(* IEC 61131-3 sources: volt/packages/volt-lsp-iec/test-corpus/lenze-mid/Device/Plc Logic/Application/Library Manager/L_IMHP_ModuleHandler, 81 files *)

(* ---- L_IMHP_COMPONENTTYPE.dut ---- *)
TYPE L_IMHP_COMPONENTTYPE :
(
	DEVICE := 101,
	IEC_RUNTIME := 102,
	LINUX_RUNTIME := 103,
	FAST_UI_RUNTIME := 104,
	FRAMEWORKSERVICE := 105,
	DEVICEFEATURES := 106,
	ETHERCATSLAVE := 201,
	ETHERCATMASTER := 202,
	FIELDBUSSLAVE := 203,
	FIELDBUSMASTER := 204,
	ETHERNET := 205,
	OPC_UA_CLIENT := 206,
	OPC_UA_SERVER := 207,
	UI_CLIENT := 208,
	UI_SERVER := 209,
	SINGLEAXISKINEMATICS := 301,
	SINGLEAXISKINEMATIK := 301,
	ROBOTKINEMATICS := 302,
	ROBOTKINEMATIC := 302,
	LOGICAXIS := 401,
	MOTIONAXIS := 402,
	VIRTUALAXIS := 403,
	ENCODERAXIS := 404,
	VIRTUALENCODERAXIS := 405,
	TECHNOLOGYFUNCTIONS := 500,
	TECHNOLOGYMODULE := 501,
	TECHNOLOGYAPPLICATION := 503,
	MACHINEMODULE := 504,
	MOTIONBASE := 505,
	COORDINATEDMOTION := 506,
	GENERALMACHINEMODULE := 551,
	GENERALAPPLICATIONMODULE := 552,
	DATAMANAGEMENT := 601,
	CLOUDCONNECTIVITY := 602,
	DATAANALYTICS := 603
);
END_TYPE

(* ---- L_IMHP_EM_CLEARERRORDATA.dut ---- *)
TYPE L_IMHP_EM_CLEARERRORDATA :
STRUCT
	VERSION : UDINT := 1;
	WERRORID : WORD;
	WTEXTREFID : WORD;
END_STRUCT
END_TYPE

(* ---- L_IMHP_EM_COMMAND.dut ---- *)
TYPE L_IMHP_EM_COMMAND :
(
	NOCOMMAND := 0,
	NOTIFYERROR := 1,
	NOTIFYERRORSHORT := 2,
	CLEARERROR := 3,
	RESETERROR := 4
);
END_TYPE

(* ---- L_IMHP_EM_EVENTPARAMETERS.dut ---- *)
TYPE L_IMHP_EM_EVENTPARAMETERS :
STRUCT
	EVENTPARAMETERS : ARRAY [1..10] OF L_IMHP_EM_ParameterItem;
END_STRUCT
END_TYPE

(* ---- L_IMHP_EM_EVENTPARAMETERSSHORT.dut ---- *)
TYPE L_IMHP_EM_EVENTPARAMETERSSHORT :
STRUCT
	EVENTPARAMETERS : ARRAY [1..10] OF L_IMHP_EM_ParameterItemShort;
END_STRUCT
END_TYPE

(* ---- L_IMHP_EM_NOTIFYERRORDATA.dut ---- *)
TYPE L_IMHP_EM_NOTIFYERRORDATA :
STRUCT
	VERSION : UDINT := 1;
	WERRORID : WORD;
	WTEXTREFID : WORD;
	SEVERITY : USINT;
	PRIORITY : USINT;
	GROUP : USINT;
END_STRUCT
END_TYPE

(* ---- L_IMHP_EM_PARAMETERITEM.dut ---- *)
TYPE L_IMHP_EM_PARAMETERITEM :
STRUCT
	SIZE : BYTE;
	ETYPE : INT;
	VALUE : L_IMHP_EM_ParaValue;
END_STRUCT
END_TYPE

(* ---- L_IMHP_EM_PARAMETERITEMSHORT.dut ---- *)
TYPE L_IMHP_EM_PARAMETERITEMSHORT :
STRUCT
	SIZE : BYTE;
	ETYPE : INT;
	VALUE : L_IMHP_EM_ParaValueShort;
END_STRUCT
END_TYPE

(* ---- L_IMHP_EM_PARAVALUE.dut ---- *)
TYPE L_IMHP_EM_PARAVALUE :
UNION
	DWVALUE : DWORD;
	DNVALUE : DINT;
	FVALUE : REAL;
	STVALUE : STRING;
	DWTEXTLISTID : DWORD;
END_UNION
END_TYPE

(* ---- L_IMHP_EM_PARAVALUESHORT.dut ---- *)
TYPE L_IMHP_EM_PARAVALUESHORT :
UNION
	DWVALUE : DWORD;
	DNVALUE : DINT;
	RVALUE : REAL;
	LRVALUE : LREAL;
	DWTEXTLISTID : DWORD;
END_UNION
END_TYPE

(* ---- L_IMHP_EM_REGISTERDATA.dut ---- *)
TYPE L_IMHP_EM_REGISTERDATA :
STRUCT
	VERSION : UDINT := 1;
	CMPNAME : POINTER TO STRING;
	LAYER : BYTE;
	TEXTREFID : WORD;
	ADDITIONALCMPINFOS : DWORD;
END_STRUCT
END_TYPE

(* ---- L_IMHP_EM_SERVERITYLEVEL.dut ---- *)
TYPE L_IMHP_EM_SERVERITYLEVEL :
(
	NO_RESPONSE := 0,
	FAULT_CIA402 := 1,
	WARNING := 2,
	INFORMATION := 11,
	WARNING_LOCK := 13,
	TROUBLE_LOG := 15,
	TROUBLE := 16,
	FAULT_LOG := 18,
	FAULT_FAST_STOP := 19,
	FAULT_QSP := 20,
	FAULT_QSP_CINH := 21,
	FAULT := 23
);
END_TYPE

(* ---- L_IMHP_LAYER.dut ---- *)
TYPE L_IMHP_LAYER :
(
	BASE_SETTINGS := 4,
	COMMUNICATION := 5,
	KINEMATICS := 6,
	MOTION := 7,
	TECH_APPLICATION := 8,
	PROCESS_CONTROL := 9
);
END_TYPE

(* ---- L_IMHP_LM_APPLICATIONCREDITCONFIGURATION.dut ---- *)
TYPE L_IMHP_LM_APPLICATIONCREDITCONFIGURATION :
STRUCT
	VERSION : DWORD := 1;
	SIZE : DWORD := SIZEOF(L_IMHP_LM_ApplicationCreditConfiguration);
	FAST_TOOLBOX : DWORD := 0;
	FAST_SERVICES : DWORD := 0;
	FAST_UI : DWORD := 0;
	OPC_UA : DWORD := 0;
	DEVICE_FEATURES : DWORD := 0;
	ADDITIONAL_BUDGETS : ARRAY [0..14] OF DWORD := [0, 0, 0, 0, 0, 0, 0, 0, 0, 0, 0, 0, 0, 0, 0];
END_STRUCT
END_TYPE

(* ---- L_IMHP_LM_APPLICATIONCREDITINFO.dut ---- *)
TYPE L_IMHP_LM_APPLICATIONCREDITINFO :
STRUCT
	VERSION : DWORD := 1;
	SIZE : DWORD := SIZEOF(L_IMHP_LM_ApplicationCreditInfo);
	AVAILABLEAPPLICATIONCREDIT : DWORD := 0;
	MAXAPPLICATIONCREDIT : DWORD := 0;
	USEDAPPLICATIONCREDIT : DWORD := 0;
END_STRUCT
END_TYPE

(* ---- L_IMHP_LM_BLISTDATA.dut ---- *)
TYPE L_IMHP_LM_BLISTDATA :
STRUCT
	VERSION : DWORD := 1;
	SIZE : DWORD := SIZEOF(L_IMHP_LM_BListData);
	COMPONENTNAME : POINTER TO STRING := 0;
	INSTANCEPATH : POINTER TO STRING := 0;
END_STRUCT
END_TYPE

(* ---- L_IMHP_LM_COMMAND.dut ---- *)
TYPE L_IMHP_LM_COMMAND :
(
	NOCOMMAND := 0,
	WRITECOMPONENTLIST := 1,
	GETAPPCREDITOFCOMPONENT := 2,
	GETAPPCREDITINFO := 3,
	ACTIVATEAPPCREDIT := 4,
	GETMODIFICATIONTIME := 5
);
END_TYPE

(* ---- L_IMHP_LM_CONFIGMODEDATA.dut ---- *)
TYPE L_IMHP_LM_CONFIGMODEDATA :
STRUCT
	VERSION : DWORD := 1;
	SIZE : DWORD := SIZEOF(L_IMHP_LM_ConfigModeData);
	UDICONFIGMODE : UDINT := 0;
END_STRUCT
END_TYPE

(* ---- L_IMHP_LM_CONFIGURECOMMAND.dut ---- *)
TYPE L_IMHP_LM_CONFIGURECOMMAND :
(
	NOCOMMAND := 0,
	APPCREDITCONFIGURATION := 1,
	SETCONFIGMODE := 2,
	STARTONLINECHANGEHANDLING := 3,
	FINISHONLINECHANGEHANDLING := 4
);
END_TYPE

(* ---- L_IMHP_LM_LICENSCLASS.dut ---- *)
TYPE L_IMHP_LM_LICENSCLASS :
(
	T := 1,
	F := 2,
	I := 3
);
END_TYPE

(* ---- L_IMHP_LM_REGISTERDATA.dut ---- *)
TYPE L_IMHP_LM_REGISTERDATA :
STRUCT
	VERSION : DWORD := 1;
	SIZE : DWORD := SIZEOF(L_IMHP_LM_RegisterData);
	APPLICATIONCREDIT : DWORD := 0;
	LICENSECLASS : DWORD := 0;
	LICENSECLASSNUMBER : DWORD := 0;
END_STRUCT
END_TYPE

(* ---- L_IMHP_MH_COMMAND.dut ---- *)
TYPE L_IMHP_MH_COMMAND :
(
	UPDATEACTIVESTATUS := 0,
	UPDATECOMMUNICATIONADRESS := 1,
	UPDATEPARENTCHILDRELATION := 2,
	UPDATECOMPONENTTYPE := 3,
	UPDATECOMPONENTNAME := 4
);
END_TYPE

(* ---- L_IMHP_MODULEINFO.dut ---- *)
TYPE L_IMHP_MODULEINFO :
STRUCT
	DWID : DWORD;
	SNAME : STRING;
	SPATH : STRING(255);
	SCOMMPATH : STRING(199);
	ELAYER : L_IMHP_Layer := L_IMHP_Layer.Tech_Application;
	ECOMPTYPE : L_IMHP_ComponentType := L_IMHP_ComponentType.GeneralApplicationModule;
	ESUBCOMPTYPE : DWORD;
	XCOMPACTIVE : BOOL;
	WCHILDCOUNT : WORD;
	WTEXTREFID : WORD;
	XUSELEM : BOOL;
	XUSELLM : BOOL;
	RELATIONSHIPID : L_IMHP_RelationshipID := L_IMHP_RelationshipID.ApplicationView;
	PARENTMODULE : L_IMHP_IModuleHandler;
END_STRUCT
END_TYPE

(* ---- L_IMHP_RELATIONSHIPDATA.dut ---- *)
TYPE L_IMHP_RELATIONSHIPDATA :
STRUCT
	VERSION : UDINT := 1;
	SIZE : UDINT := SIZEOF(L_IMHP_RelationshipData);
	RELATIONSHIPID : L_IMHP_RelationshipID;
	PARENTHANDLE : RTS_IEC_HANDLE;
END_STRUCT
END_TYPE

(* ---- L_IMHP_RELATIONSHIPID.dut ---- *)
TYPE L_IMHP_RELATIONSHIPID :
(
	NORELATIONSHIP := 0,
	APPLICATIONVIEW := 1,
	COMMUNICATIONVIEW := 2,
	ASSETVIEW := 3
);
END_TYPE

(* ---- L_IMHP_REQUESTEDSERVICE.dut ---- *)
TYPE L_IMHP_REQUESTEDSERVICE :
STRUCT
	VERSION : UDINT := 1;
	SIZE : UDINT := SIZEOF(L_IMHP_RequestedService);
	SERVICEID : L_IMHP_ServiceID;
	SIZEOFREGISTRATIONDATA : UDINT;
	PREGISTRATIONDATA : POINTER TO BYTE;
	SERVICEAVAILABLE : UDINT;
	SERVICEVERSION : UDINT;
	REGISTRATIONSTATUS : UDINT;
	SIZEOFRESULTDATA : UDINT;
	PRESULTDATA : POINTER TO BYTE;
END_STRUCT
END_TYPE

(* ---- L_IMHP_SERVICEAVAILABLEDATA.dut ---- *)
TYPE L_IMHP_SERVICEAVAILABLEDATA :
STRUCT
	VERSION : UDINT := 1;
	SIZE : UDINT := SIZEOF(L_IMHP_ServiceAvailableData);
	SERVICEID : L_IMHP_ServiceID;
	SERVICEAVAILABLE : UDINT;
	SERVICEVERSION : UDINT;
END_STRUCT
END_TYPE

(* ---- L_IMHP_SERVICEID.dut ---- *)
TYPE L_IMHP_SERVICEID :
(
	NOSERVICE := 0,
	LENZEMODULEHANDLER := 1,
	LENZEERRORMANAGEMENT := 2,
	LENZESTATEHANDLER := 3,
	LENZELICENSEMANAGER := 4,
	LENZEASSETMANAGER := 5
);
END_TYPE

(* ---- L_IMHP_CONSTANTS.gvl ---- *)
VAR_GLOBAL
	GC_MAXCOMPIDX : WORD := 100;
END_VAR

(* ---- L_IMHP_INTERN.gvl ---- *)
VAR_GLOBAL
	XERRORHANDLINGFORI950 : BOOL;
	DEVICEMODULEHANDLER : L_IMHP_DeviceModule;
	COMPONENTREGISTRATION : L_IMHP_HandleComponentRegistration;
END_VAR

(* ---- L_IMHP_IFASTFRAMECONFIG.itf ---- *)
INTERFACE L_IMHP_IFASTFRAMECONFIG
END_INTERFACE

METHOD ADDPARAMETERINTERFACE
VAR_INPUT
	IIODRVPARAMETER : ICmpIoDrvParameter;
END_VAR
END_METHOD

(* ---- L_IMHP_IMODULEHANDLER.itf ---- *)
INTERFACE L_IMHP_IMODULEHANDLER
END_INTERFACE

METHOD ACTIVATEAPPCREDITS : BOOL
VAR_INPUT
	XACTIVATE : BOOL;
END_VAR
END_METHOD

METHOD ADDAPPCREDIT
VAR_INPUT
	CREDIT : UDINT;
END_VAR
END_METHOD

METHOD CHECKERRORRESETOCCURED : BOOL
VAR_IN_OUT
	RESETTIME : SYSTIME;
END_VAR
END_METHOD

METHOD CHECKERRORRESETTRIGGER : BOOL
VAR_IN_OUT
	LASTTRIGGERTIME : TIME;
END_VAR
END_METHOD

METHOD CLEARSEVERITYANDREACTION
VAR_INPUT
	ESEVERITY : USINT;
	DISEVERITYCOUNT : DINT;
	EREACTION : WORD;
	DIREACTIONCOUNT : DINT;
	XHANDLEASFORWARDEDSEVERITY : BOOL;
END_VAR
END_METHOD

METHOD FORWARDLOGENTRYCLEAR
VAR_INPUT
	WERRORID : WORD;
	WTEXTREFID : WORD;
END_VAR
END_METHOD

METHOD FORWARDLOGENTRYNOTIFY
VAR_INPUT
	WERRORID : WORD;
	WTEXTREFID : WORD;
	SEVERITY : USINT;
	REACTION : UINT;
	PRIORITY : USINT;
	GROUP : USINT;
END_VAR
END_METHOD

METHOD FORWARDSEVERITYSUBMODULES
VAR_INPUT
	XENABLE : BOOL;
END_VAR
END_METHOD

METHOD GETSEVERITY
VAR_INPUT
	XINCLUDECHILDREN : BOOL;
	XDISABLESUBMODULES : BOOL;
	XINCLUDEOWNMODULE : BOOL;
	XINCLUDEEXTMODULE : BOOL;
	PSEVERITYSTATUS : POINTER TO BYTE;
	PREACTIONSTATUS : POINTER TO BYTE;
END_VAR
VAR_OUTPUT
	EHIGHESTSEVERITY : USINT;
	EHIGHESTREACTION : WORD;
	AFFECTEDMODULE : L_IMHP_IModuleHandler;
END_VAR
END_METHOD

METHOD GETSEVERITY2
VAR_INPUT
	XINCLUDECHILDREN : BOOL;
	XDISABLESUBMODULES : BOOL := FALSE;
	XDISABLEINTERNALCHILDS : BOOL := FALSE;
	XINCLUDEOWNMODULE : BOOL := TRUE;
	XINCLUDEEXTMODULE : BOOL := TRUE;
	PSEVERITYSTATUS : POINTER TO BYTE;
	PREACTIONSTATUS : POINTER TO BYTE;
END_VAR
VAR_OUTPUT
	EHIGHESTSEVERITY : USINT;
	EHIGHESTREACTION : WORD;
	AFFECTEDMODULE : L_IMHP_IModuleHandler;
END_VAR
END_METHOD

METHOD GETSEVERITYCHILD
VAR_INPUT
	WCHILD : WORD;
END_VAR
VAR_OUTPUT
	EHIGHESTSEVERITY : USINT;
	EHIGHESTREACTION : WORD;
	AFFECTEDMODULE : L_IMHP_IModuleHandler;
END_VAR
END_METHOD

METHOD READACTUALERRORCODE
VAR_OUTPUT
	ESEVERITY : USINT;
	EREACTION : WORD;
	DWERRORCODE : DWORD;
END_VAR
END_METHOD

METHOD RESETCHILDERROR
END_METHOD

METHOD RESETCHILDERROR2
VAR_INPUT
	PERRORLIST : POINTER TO RTS_IEC_HANDLE;
	PWCOUNT : POINTER TO WORD;
	MAXCOUNT : WORD;
END_VAR
END_METHOD

METHOD SETERRORRESETTRIGGER
END_METHOD

METHOD SETPARENT
VAR_INPUT
	MODULEHANDLERPARENT : L_IMHP_IModuleHandler;
	RELATIONSHIP : L_IMHP_RelationshipID := L_IMHP_RelationshipID.ApplicationView;
END_VAR
END_METHOD

METHOD SYNCSEVERITYANDREACTIONCOUNTER
VAR_INPUT
	XHANDLEASFORWARDEDSEVERITY : BOOL;
END_VAR
VAR_IN_OUT
	SEVERITYCOUNTER_CHILD : L_IE1P_SeverityCounter;
	REACTIONCOUNTER_CHILD : L_IE1P_ReactionCounter;
	REACTIONCOUNTERWARNING_CHILD : L_IE1P_ReactionCounter;
	REACTIONCOUNTERINFORMATION_CHILD : L_IE1P_ReactionCounter;
	REACTIONCOUNTERWARNINGLOCK_CHILD : L_IE1P_ReactionCounter;
	REACTIONCOUNTERFAULTLOG_CHILD : L_IE1P_ReactionCounter;
	REACTIONCOUNTERFAULT_CHILD : L_IE1P_ReactionCounter;
END_VAR
END_METHOD

METHOD UPDATEACTIVESTATUS
VAR_INPUT
	XACTIVE : BOOL;
END_VAR
END_METHOD

METHOD UPDATESEVERITYANDREACTION
VAR_INPUT
	ESEVERITY : USINT;
	EREACTION : WORD;
	XHANDLEASFORWARDEDSEVERITY : BOOL;
END_VAR
END_METHOD

METHOD ADDCHILD
VAR_INPUT
	MODULEHANDLERCHILD : L_IMHP_IModuleHandler;
	RELATIONSHIP : L_IMHP_RelationshipID := L_IMHP_RelationshipID.ApplicationView;
END_VAR
END_METHOD

METHOD GETCHILD : L_IMHP_IModuleHandler
VAR_INPUT
	WNBR : WORD;
END_VAR
END_METHOD

METHOD REMOVECHILD
VAR_INPUT
	MODULEHANDLERCHILD : L_IMHP_IModuleHandler;
END_VAR
END_METHOD

METHOD SETCHILDFORDELAYEDREGISTRATION
VAR_INPUT
	MODULEHANDLERCHILD : L_IMHP_IModuleHandler;
	RELATIONSHIP : L_IMHP_RelationshipID := L_IMHP_RelationshipID.ApplicationView;
END_VAR
END_METHOD

METHOD GETCOMMPATH
VAR_IN_OUT
	SCOMMPATH : STRING(199);
END_VAR
END_METHOD

METHOD GETCOMPTYPE : L_IMHP_ComponentType
END_METHOD

METHOD GETDEVICECONNECTOR : POINTER TO IoConfigConnector
END_METHOD

METHOD GETMODULEINFO : BOOL
VAR_IN_OUT
	MODULEINFO : L_IMHP_ModuleInfo;
END_VAR
END_METHOD

METHOD GETMODULENAME
VAR_IN_OUT
	SNAME : STRING;
END_VAR
END_METHOD

METHOD REGISTEREDONSERVICE : BOOL
VAR_INPUT
	SERVICEID : L_IMHP_ServiceID;
END_VAR
END_METHOD

(* ---- L_IMHP_IREGISTERCOMPONENT.itf ---- *)
INTERFACE L_IMHP_IREGISTERCOMPONENT
END_INTERFACE

METHOD DOREGISTER
END_METHOD

METHOD UPDATEDEPENDENCIES
END_METHOD

(* ---- GETBOOLEANPROPERTY.pou ---- *)
FUNCTION GETBOOLEANPROPERTY : BOOL
VAR_INPUT
	STKEY : WSTRING;
END_VAR
END_FUNCTION

(* ---- GETCOMPANY.pou ---- *)
FUNCTION GETCOMPANY : WSTRING
END_FUNCTION

(* ---- GETNUMBERPROPERTY.pou ---- *)
FUNCTION GETNUMBERPROPERTY : DINT
VAR_INPUT
	STKEY : WSTRING;
END_VAR
END_FUNCTION

(* ---- GETTEXTPROPERTY.pou ---- *)
FUNCTION GETTEXTPROPERTY : WSTRING
VAR_INPUT
	STKEY : WSTRING;
END_VAR
END_FUNCTION

(* ---- GETTEXTPROPERTY2.pou ---- *)
FUNCTION GETTEXTPROPERTY2 : POINTER TO WSTRING
VAR_INPUT
	STKEY : WSTRING;
END_VAR
END_FUNCTION

(* ---- GETTITLE.pou ---- *)
FUNCTION GETTITLE : WSTRING
END_FUNCTION

(* ---- GETVERSION.pou ---- *)
FUNCTION GETVERSION : VERSION
END_FUNCTION

(* ---- GETVERSIONPROPERTY.pou ---- *)
FUNCTION GETVERSIONPROPERTY : VERSION
VAR_INPUT
	STKEY : WSTRING;
END_VAR
END_FUNCTION

(* ---- L_IHMP_SIMPLEREGISTERCOMPONENTFORLEM.pou ---- *)
FUNCTION L_IHMP_SIMPLEREGISTERCOMPONENTFORLEM : BOOL
VAR_INPUT
	SCOMPNAME : STRING;
	SPATH : STRING(255);
	UILAYER : UINT;
	UDICOMPTYPE : UDINT;
	UITEXTREFID : UINT;
	UIREAKTIONITF : UINT;
END_VAR
VAR_OUTPUT
	REGISTERDLEMHANDLE : RTS_IEC_HANDLE;
	REGISTERDLMHHANDLE : RTS_IEC_HANDLE;
END_VAR
END_FUNCTION

(* ---- L_IHMP_SIMPLEREGISTERCOMPONENTFORLLM.pou ---- *)
FUNCTION L_IHMP_SIMPLEREGISTERCOMPONENTFORLLM : RTS_IEC_HANDLE
VAR_INPUT
	SCOMPNAME : STRING;
	SPATH : STRING(255);
	UILAYER : UINT;
	UDICOMPTYPE : UDINT;
	UDICOMPSUBTYPE : UDINT;
	DWAPPLICATIONCREDIT : DWORD := 0;
	DWLICENSECLASS : L_IMHP_LM_LicensClass := 0;
	DWLICENSECLASSNUMBER : DWORD := 0;
END_VAR
END_FUNCTION

(* ---- L_IMHP_ADDREACTIONCOUNTER.pou ---- *)
FUNCTION L_IMHP_ADDREACTIONCOUNTER : BOOL
VAR_IN_OUT
	REACTIONCOUNTERIN1 : L_IE1P_ReactionCounter;
	REACTIONCOUNTERIN2 : L_IE1P_ReactionCounter;
	REACTIONCOUNTEROUT : L_IE1P_ReactionCounter;
END_VAR
END_FUNCTION

(* ---- L_IMHP_ADDSEVERITYCOUNTER.pou ---- *)
FUNCTION L_IMHP_ADDSEVERITYCOUNTER : BOOL
VAR_IN_OUT
	SEVERITYCOUNTERIN1 : L_IE1P_SeverityCounter;
	SEVERITYCOUNTERIN2 : L_IE1P_SeverityCounter;
	SEVERITYCOUNTEROUT : L_IE1P_SeverityCounter;
END_VAR
END_FUNCTION

(* ---- L_IMHP_CALLCYCLICFUNCTIONS.pou ---- *)
FUNCTION L_IMHP_CALLCYCLICFUNCTIONS : BOOL
END_FUNCTION

(* ---- L_IMHP_EM_CLEARERROR.pou ---- *)
FUNCTION L_IMHP_EM_CLEARERROR : UDINT
VAR_INPUT
	ERRORHANDLERID : RTS_IEC_HANDLE;
	WERRORID : WORD;
	WTEXTREFID : WORD;
END_VAR
END_FUNCTION

(* ---- L_IMHP_EM_NOTIFYERROR.pou ---- *)
FUNCTION L_IMHP_EM_NOTIFYERROR : UDINT
VAR_INPUT
	ERRORHANDLERID : RTS_IEC_HANDLE;
	WERRORID : WORD;
	WTEXTREFID : WORD;
	SEVERITY : USINT;
	PRIORITY : USINT;
	GROUP : USINT;
	XNOLOGENTRY : BOOL := FALSE;
END_VAR
END_FUNCTION

(* ---- L_IMHP_EM_NOTIFYERRORNOLOGBOOK.pou ---- *)
FUNCTION L_IMHP_EM_NOTIFYERRORNOLOGBOOK : UDINT
VAR_INPUT
	ERRORHANDLERID : RTS_IEC_HANDLE;
	WERRORID : WORD;
	WTEXTREFID : WORD;
	SEVERITY : USINT;
	REACTION : UINT;
	PRIORITY : USINT;
	GROUP : USINT;
END_VAR
END_FUNCTION

(* ---- L_IMHP_EM_NOTIFYERRORWITHPAR.pou ---- *)
FUNCTION L_IMHP_EM_NOTIFYERRORWITHPAR : UDINT
VAR_INPUT
	ERRORHANDLERID : RTS_IEC_HANDLE;
	WERRORID : WORD;
	WTEXTREFID : WORD;
	SEVERITY : USINT;
	PRIORITY : USINT;
	GROUP : USINT;
	XNOLOGENTRY : BOOL := FALSE;
	PARCOUNT : UINT;
	PPAR : POINTER TO L_IMHP_EM_ParameterItemShort;
END_VAR
END_FUNCTION

(* ---- L_IMHP_EM_RESETERROR.pou ---- *)
FUNCTION L_IMHP_EM_RESETERROR : UDINT
VAR_INPUT
	ERRORHANDLERID : RTS_IEC_HANDLE;
END_VAR
END_FUNCTION

(* ---- L_IMHP_EM_RESETERRORGLOBAL.pou ---- *)
FUNCTION L_IMHP_EM_RESETERRORGLOBAL : UDINT
VAR_INPUT
	ERRORHANDLERID : RTS_IEC_HANDLE;
END_VAR
END_FUNCTION

(* ---- L_IMHP_EM_RESETERRORLIST.pou ---- *)
FUNCTION L_IMHP_EM_RESETERRORLIST : UDINT
VAR_INPUT
	PERRORLIST : POINTER TO RTS_IEC_HANDLE;
	WCOUNT : WORD;
END_VAR
END_FUNCTION

(* ---- L_IMHP_GETCOMPNAMEBYINSTANCEID.pou ---- *)
FUNCTION L_IMHP_GETCOMPNAMEBYINSTANCEID : STRING
VAR_INPUT
	MODULEINSTANCEID : DWORD;
END_VAR
VAR_OUTPUT
	EERRORID : L_IE1P_Error;
END_VAR
END_FUNCTION

(* ---- L_IMHP_GETDEVICEMODULEHANDLER.pou ---- *)
FUNCTION L_IMHP_GETDEVICEMODULEHANDLER : L_IMHP_IModuleHandler
END_FUNCTION

(* ---- L_IMHP_GETHIGHESTREACTION.pou ---- *)
FUNCTION L_IMHP_GETHIGHESTREACTION : BOOL
VAR_INPUT
	EREACTION1 : L_IE1P_Reaction;
	MODULEHANDLER1 : POINTER TO BYTE;
	EREACTION2 : L_IE1P_Reaction;
	MODULEHANDLER2 : POINTER TO BYTE;
END_VAR
VAR_OUTPUT
	EREACTION : L_IE1P_Reaction;
	MODULEHANDLER : POINTER TO BYTE;
END_VAR
END_FUNCTION

(* ---- L_IMHP_GETHIGHESTSEVERITYANDREACTION.pou ---- *)
FUNCTION L_IMHP_GETHIGHESTSEVERITYANDREACTION : BOOL
VAR_INPUT
	ESEVERITY1 : L_IE1P_SeverityLevel;
	EREACTION1 : L_IE1P_Reaction;
	MODULEHANDLER1 : POINTER TO BYTE;
	ESEVERITY2 : L_IE1P_SeverityLevel;
	EREACTION2 : L_IE1P_Reaction;
	MODULEHANDLER2 : POINTER TO BYTE;
END_VAR
VAR_OUTPUT
	ESEVERITY : L_IE1P_SeverityLevel;
	EREACTION : L_IE1P_Reaction;
	MODULEHANDLER : POINTER TO BYTE;
END_VAR
END_FUNCTION

(* ---- L_IMHP_GETLAYERFROMCOMPTYPE.pou ---- *)
FUNCTION L_IMHP_GETLAYERFROMCOMPTYPE : L_IMHP_Layer
VAR_INPUT
	ECOMPTYPE : L_IMHP_ComponentType;
END_VAR
END_FUNCTION

(* ---- L_IMHP_HANDLELMF1CLASSES.pou ---- *)
FUNCTION L_IMHP_HANDLELMF1CLASSES : RTS_IEC_HANDLE
VAR_INPUT
	MODE : WORD;
	SCOMPNAME : STRING;
	SPATH : STRING(255);
	UILAYER : UINT;
	UDICOMPTYPE : UDINT;
	UDICOMPSUBTYPE : UDINT;
	DWAPPLICATIONCREDIT : DWORD := 0;
	DWLICENSECLASS : L_IMHP_LM_LicensClass := 0;
	DWLICENSECLASSNUMBER : DWORD := 0;
END_VAR
END_FUNCTION

(* ---- L_IMHP_HANDLELMF2CLASSES.pou ---- *)
FUNCTION L_IMHP_HANDLELMF2CLASSES : RTS_IEC_HANDLE
VAR_INPUT
	MODE : WORD;
	SCOMPNAME : STRING;
	SPATH : STRING(255);
	UILAYER : UINT;
	UDICOMPTYPE : UDINT;
	UDICOMPSUBTYPE : UDINT;
	DWAPPLICATIONCREDIT : DWORD := 0;
	DWLICENSECLASS : L_IMHP_LM_LicensClass := 0;
	DWLICENSECLASSNUMBER : DWORD := 0;
END_VAR
END_FUNCTION

(* ---- L_IMHP_HANDLEREGISTRATIONAFTERONLINECHANGE.pou ---- *)
FUNCTION L_IMHP_HANDLEREGISTRATIONAFTERONLINECHANGE : BOOL
VAR_INPUT
	ITFREGISTERCOMPONENT : L_IMHP_IRegisterComponent;
END_VAR
END_FUNCTION

(* ---- L_IMHP_ISSERVICEAVAILABLE.pou ---- *)
FUNCTION L_IMHP_ISSERVICEAVAILABLE : BOOL
VAR_INPUT
	SERVICE : L_IMHP_ServiceID;
END_VAR
END_FUNCTION

(* ---- L_IMHP_ISSERVICEAVAILABLELLM.pou ---- *)
FUNCTION L_IMHP_ISSERVICEAVAILABLELLM : BOOL
END_FUNCTION

(* ---- L_IMHP_LM_ACTIVATEAPPCREDITS.pou ---- *)
FUNCTION L_IMHP_LM_ACTIVATEAPPCREDITS : BOOL
VAR_INPUT
	MODULEHANDLERID : RTS_IEC_HANDLE;
	XACTIVATE : BOOL;
END_VAR
END_FUNCTION

(* ---- L_IMHP_LM_CHECKLICENSESTRING.pou ---- *)
FUNCTION L_IMHP_LM_CHECKLICENSESTRING : BOOL
VAR_INPUT
	SLICINFO : STRING;
END_VAR
VAR_IN_OUT
	UDIAPPLICATIONCREDIT : DWORD;
	ELICENSECLASS : L_IMHP_LM_LicensClass;
	UDILICENSECLASSNUMBER : DWORD;
END_VAR
END_FUNCTION

(* ---- L_IMHP_LM_GETAPPCREDITINFO.pou ---- *)
FUNCTION L_IMHP_LM_GETAPPCREDITINFO : BOOL
VAR_INPUT
	MODULEHANDLERID : RTS_IEC_HANDLE;
	PAPPCREDITINFO : POINTER TO L_IMHP_LM_ApplicationCreditInfo;
END_VAR
END_FUNCTION

(* ---- L_IMHP_LM_SETAPPCREDITCONFIGMODE.pou ---- *)
FUNCTION L_IMHP_LM_SETAPPCREDITCONFIGMODE : BOOL
VAR_INPUT
	DWAPPCREDITCONFIGMODE : UDINT;
END_VAR
END_FUNCTION

(* ---- L_IMHP_LM_SETAPPCREDITCONFIGURATION.pou ---- *)
FUNCTION L_IMHP_LM_SETAPPCREDITCONFIGURATION : BOOL
VAR_INPUT
	PAPPCREDITCONFIG : POINTER TO L_IMHP_LM_ApplicationCreditConfiguration;
END_VAR
END_FUNCTION

(* ---- L_IMHP_MODULEREGISTRATIONAFTERONLINECHANGESUPPORTED.pou ---- *)
FUNCTION L_IMHP_MODULEREGISTRATIONAFTERONLINECHANGESUPPORTED : BOOL
END_FUNCTION

(* ---- L_IMHP_READERRORDATAFROMCOMPONENTLIST.pou ---- *)
FUNCTION L_IMHP_READERRORDATAFROMCOMPONENTLIST : BOOL
VAR_INPUT
	MODULEHANDLE : UDINT;
	PDATA : POINTER TO L_IE1P_Types.L_IE1P_ReadErrorData;
END_VAR
VAR_OUTPUT
	SEVERITY : L_IE1P_SeverityLevel;
	ERRORCODE : DWORD := 0;
END_VAR
VAR_IN_OUT
	DWCOMPIDX : DWORD;
END_VAR
END_FUNCTION

(* ---- L_IMHP_REGISTRATIONAFTERONLINECHANGEBUSY.pou ---- *)
FUNCTION L_IMHP_REGISTRATIONAFTERONLINECHANGEBUSY : BOOL
END_FUNCTION

(* ---- GLOBALTEXTLIST.pou ---- *)
FUNCTION_BLOCK GLOBALTEXTLIST
VAR
	M_TEXTLISTFILE : STRING(255);
	_STNAMESPACE : STRING;
END_VAR
END_FUNCTION_BLOCK

(* ---- L_IMHP_DEVICEMODULE.pou ---- *)
FUNCTION_BLOCK L_IMHP_DEVICEMODULE EXTENDS L_IMHP_ModuleHandler
VAR
	COMPNAME : STRING;
	ERRORHANDLE : RTS_IEC_HANDLE;
	FORWARDLOGENTRYENABLED : BOOL;
	FORWARDSEVERITYTOPARENT : BOOL;
	GETMODULEHANDLERFB : POINTER TO BYTE;
	MODULEHANDLE : RTS_IEC_HANDLE;
	REGISTRATIONBUSY : BOOL;
END_VAR
END_FUNCTION_BLOCK

METHOD GETAPPNAME
END_METHOD

METHOD FB_INIT : BOOL
VAR_INPUT
	BINITRETAINS : BOOL;
	BINCOPYCODE : BOOL;
END_VAR
END_METHOD

METHOD ACTIVATEAPPCREDITS : BOOL
VAR_INPUT
	XACTIVATE : BOOL;
END_VAR
END_METHOD

METHOD ADDCHILD
VAR_INPUT
	MODULEHANDLERCHILD : L_IMHP_IModuleHandler;
	RELATIONSHIP : L_IMHP_RelationshipID := L_IMHP_RelationshipID.ApplicationView;
END_VAR
END_METHOD

METHOD REMOVECHILD
VAR_INPUT
	MODULEHANDLERCHILD : L_IMHP_IModuleHandler;
END_VAR
END_METHOD

METHOD RESETCHILDERROR
END_METHOD

METHOD RESETCHILDERROR2
VAR_INPUT
	PERRORLIST : POINTER TO RTS_IEC_HANDLE;
	PWCOUNT : POINTER TO WORD;
	MAXCOUNT : WORD;
END_VAR
END_METHOD

METHOD SETPARENT
VAR_INPUT
	MODULEHANDLERPARENT : L_IMHP_IModuleHandler;
	RELATIONSHIP : L_IMHP_RelationshipID := L_IMHP_RelationshipID.ApplicationView;
END_VAR
END_METHOD

METHOD UPDATEACTIVESTATUS
VAR_INPUT
	XACTIVE : BOOL;
END_VAR
END_METHOD

(* ---- L_IMHP_FASTFRAMECONFIGURATION.pou ---- *)
FUNCTION_BLOCK L_IMHP_FASTFRAMECONFIGURATION EXTENDS IoDrvBase
VAR
	M_IIODRVPARAMETER : ICmpIoDrvParameter;
	M_IIODRV : ICmpIoDrv;
	M_IFASTFRAMCONFIG : L_IMHP_IFastFrameConfig;
	DWREADCALL : DWORD;
	DWWRITECALL : DWORD;
	UPDATECOUNT : WORD;
	SUBCONNECTORPARAMETERACCES : ARRAY [1..5] OF ICmpIoDrvParameter;
	COUNTSUBCONNECTORPARAMETERACCES : WORD;
END_VAR
END_FUNCTION_BLOCK

METHOD ADDPARAMETERINTERFACE
VAR_INPUT
	IIODRVPARAMETER : ICmpIoDrvParameter;
END_VAR
END_METHOD

METHOD INITIALIZE : UDINT
VAR_INPUT
	WMODULETYPE : UINT;
	DWINSTANCE : UDINT;
	PCONNECTOR : POINTER TO IoConfigConnector;
END_VAR
END_METHOD

METHOD IODRVREADPARAMETER : UDINT
VAR_INPUT
	PCONNECTOR : POINTER TO IoConfigConnector;
	PPARAMETER : POINTER TO IoConfigParameter;
	PDATA : POINTER TO BYTE;
	DWBITSIZE : DWORD;
	DWBITOFFSET : DWORD;
END_VAR
END_METHOD

METHOD IODRVUPDATECONFIGURATION : UDINT
VAR_INPUT
	PCONNECTORLIST : POINTER TO IoConfigConnector;
	NCOUNT : DINT;
END_VAR
END_METHOD

METHOD IODRVUPDATEMAPPING : UDINT
VAR_INPUT
	PTASKMAPLIST : POINTER TO IoConfigTaskMap;
	NCOUNT : DINT;
END_VAR
END_METHOD

METHOD IODRVWRITEPARAMETER : UDINT
VAR_INPUT
	PCONNECTOR : POINTER TO IoConfigConnector;
	PPARAMETER : POINTER TO IoConfigParameter;
	PDATA : POINTER TO BYTE;
	DWBITSIZE : DWORD;
	DWBITOFFSET : DWORD;
END_VAR
END_METHOD

METHOD QUERYINTERFACE : POINTER TO POINTER TO BYTE
VAR_INPUT
	IID : DWORD;
	PRESULT : POINTER TO UDINT;
END_VAR
END_METHOD

METHOD FB_INIT : BOOL
VAR_INPUT
	BINITRETAINS : BOOL;
	BINCOPYCODE : BOOL;
END_VAR
END_METHOD

(* ---- L_IMHP_GETCHILDMODULE.pou ---- *)
FUNCTION_BLOCK L_IMHP_GETCHILDMODULE
VAR_INPUT
	MODULEHANDLER : L_IMHP_IModuleHandler;
	WCHILD : WORD;
END_VAR
VAR_OUTPUT
	CHILDMODULEHANDLER : L_IMHP_IModuleHandler;
END_VAR
END_FUNCTION_BLOCK

(* ---- L_IMHP_GETMODULEINFO.pou ---- *)
FUNCTION_BLOCK L_IMHP_GETMODULEINFO
VAR_INPUT
	MODULEHANDLER : L_IMHP_IModuleHandler;
END_VAR
VAR_OUTPUT
	SNAME : STRING;
	ELAYER : L_IMHP_Layer := L_IMHP_Layer.Tech_Application;
	ECOMPTYPE : L_IMHP_ComponentType := L_IMHP_ComponentType.GeneralApplicationModule;
	XCOMPACTIVE : BOOL;
	WCHILDCOUNT : WORD;
END_VAR
VAR
	MODULEINFO : L_IMHP_ModuleInfo;
	MODULEHANDLERINT : L_IMHP_IModuleHandler;
END_VAR
END_FUNCTION_BLOCK

(* ---- L_IMHP_HANDLECOMPONENTREGISTRATION.pou ---- *)
FUNCTION_BLOCK L_IMHP_HANDLECOMPONENTREGISTRATION
VAR
	DWCALLAFTERONLINECHANGE : DWORD;
	XINFORMLMH : BOOL;
	WREGISTERCOUNT : WORD := 0;
	AITFREGISTERCOMPONENT : ARRAY [1..c_maxRegister] OF L_IMHP_IRegisterComponent;
	XREGISTRATIONBUSY : BOOL;
	XCYCLICREGISTRATIONSTART : BOOL;
	WSTARTCOUNTER : WORD := 1;
	C_MAXREGISTER : WORD := 500;
END_VAR
END_FUNCTION_BLOCK

METHOD CALLAFTERONLINECHANGE : BOOL
END_METHOD

METHOD CALLCYCLIC : BOOL
END_METHOD

METHOD CALLUPDATEDEBENDENCIES : BOOL
END_METHOD

METHOD INSERTREGISTRATIONDATA : BOOL
VAR_INPUT
	ITFREGISTERCOMPONENT : L_IMHP_IRegisterComponent;
END_VAR
END_METHOD

METHOD ABORT : UDINT
END_METHOD

METHOD EXECUTE : UDINT
END_METHOD

(* ---- L_IMHP_LLMHANDLING.pou ---- *)
FUNCTION_BLOCK L_IMHP_LLMHANDLING
VAR
	XLICENCEMANAGERAVAILABLE : BOOL := FALSE;
	HLICENCEMANAGER : RTS_IEC_HANDLE := RTS_INVALID_HANDLE;
	SINSTANCEPATHFULL : STRING(255);
	UILAYER : UINT;
	UDICOMPTYPE : UDINT;
	UDICOMPSUBTYPE : UDINT;
	DWAPPLICATIONCREDIT : DWORD := 0;
	DWLICENSECLASS : L_IMHP_LM_LicensClass := 0;
	DWLICENSECLASSNUMBER : DWORD := 0;
	XREGISTERONLLMDONE : BOOL;
	WBLCLASS : WORD;
END_VAR
END_FUNCTION_BLOCK

METHOD ACTIVATE : BOOL
VAR_INPUT
	XACTIVATE : BOOL;
END_VAR
END_METHOD

METHOD AFTERGLOBALINIT
END_METHOD

METHOD GETSTRINGS
VAR_IN_OUT
	SINSTANCEPATH : STRING(255);
	SINSTANCESTR : STRING(80);
END_VAR
END_METHOD

METHOD FB_EXIT : BOOL
VAR_INPUT
	BINCOPYCODE : BOOL;
END_VAR
END_METHOD

METHOD FB_INIT : BOOL
VAR_INPUT
	BINITRETAINS : BOOL;
	BINCOPYCODE : BOOL;
	UILAYER : UINT;
	UDICOMPTYPE : UDINT;
	UDICOMPSUBTYPE : UDINT;
	DWAPPLICATIONCREDIT : DWORD := 0;
	DWLICENSECLASS : L_IMHP_LM_LicensClass := 0;
	DWLICENSECLASSNUMBER : DWORD := 0;
END_VAR
END_METHOD

METHOD DOREGISTER
END_METHOD

METHOD UPDATEDEPENDENCIES
END_METHOD

(* ---- L_IMHP_MODULEHANDLER.pou ---- *)
FUNCTION_BLOCK L_IMHP_MODULEHANDLER
VAR_OUTPUT
	MODULEHANDLER : L_IMHP_IModuleHandler := THIS^;
END_VAR
VAR
	REGISTERCOMPONENTHANDLE : RTS_IEC_HANDLE;
	REGISTERLEMHANDLE : RTS_IEC_HANDLE;
	EM_REGISTERDATA : L_IMHP_EM_RegisterData;
	LLM_REGISTERDATA : L_IMHP_LM_RegisterData;
	SINSTANCEPATH : STRING(255);
	SINSTANCESTR : STRING(80);
	SCOMPNAME : STRING(80) := '';
	SINSTANCESTRFULL : STRING(255);
	ITFCALLBACK : CmpEventMgr.ICmpEventCallback;
	HEVENTACTUALERROR : RTS_IEC_HANDLE := SysTypes.RTS_INVALID_HANDLE;
	HINTERFACEACTUALERROR : RTS_IEC_HANDLE := SysTypes.RTS_INVALID_HANDLE;
	HEVENTRESETOCCURED : RTS_IEC_HANDLE := SysTypes.RTS_INVALID_HANDLE;
	HINTERFACERESETOCCURED : RTS_IEC_HANDLE := SysTypes.RTS_INVALID_HANDLE;
	ERRORRESETOCCUREDTIME : SysTime;
	ERRORRESETTRIGGERTIME : TIME;
	DWEVTCOUNT_RESETOCCURED : DWORD;
	DWEVTCOUNT_ERRORUPDATED : DWORD;
	DWCOMPIDXERRORUPDATED : DWORD := 0;
	DWERRORCODEMOD : ARRAY [0..1] OF DWORD;
	MYMODULEHANDLE : UDINT;
	ESEVERITYMOD : ARRAY [0..1] OF L_IE1P_SeverityLevel;
	ECOMPTYPESEND : L_IMHP_ComponentType;
	RELATIONSHIPREGISTRATIONSEND : L_IMHP_RelationshipData;
	XACTIVEERRORINFO : BOOL;
	XCOMPACTIVESEND : BOOL;
	XSUSPENDREGISTRATION : BOOL := FALSE;
	XREGISTERONLMHDONE : BOOL := FALSE;
	XREGISTERONAPPLICATIONVIEW : BOOL := TRUE;
	WCHILDCOUNT : WORD := 0;
	UDIAPPCREDIT : UDINT;
	MYDEVICECONNECTOR : POINTER TO IoConfigConnector;
	MYMODULEINFO : L_IMHP_ModuleInfo := STRUCT(xUseLEM := TRUE, xUseLLM := FALSE, xCompActive := TRUE, eLayer := L_IMHP_Layer.Tech_Application, eCompType := L_IMHP_ComponentType.GeneralMachineModule, eSubCompType := 0, RelationShipID := L_IMHP_RelationshipID.ApplicationView, ParentModule := 0, wTextRefID := 16#2C00);
	OWNMODULEHANDLER : L_IMHP_IModuleHandler;
	CHILDMODULES : ARRAY [0..maxChild] OF L_IMHP_IModuleHandler;
	CHILDSEVERITY : ARRAY [0..maxChild] OF L_IE1P_SeverityLevel;
	CHILDREACTION : ARRAY [0..maxChild] OF L_IE1P_Reaction;
	MODULEREACTIONCOUNTER : L_IE1P_ReactionCounter;
	MODULEREACTIONCOUNTERINFORMATION : L_IE1P_ReactionCounter;
	MODULEREACTIONCOUNTERWARNING : L_IE1P_ReactionCounter;
	MODULEREACTIONCOUNTERWARNINGLOCK : L_IE1P_ReactionCounter;
	MODULEREACTIONCOUNTERFAULTLOG : L_IE1P_ReactionCounter;
	MODULEREACTIONCOUNTERFAULT : L_IE1P_ReactionCounter;
	MODULESEVERITYCOUNTER : L_IE1P_SeverityCounter;
	EXTREACTIONCOUNTER : L_IE1P_ReactionCounter;
	EXTREACTIONCOUNTERINFORMATION : L_IE1P_ReactionCounter;
	EXTREACTIONCOUNTERWARNING : L_IE1P_ReactionCounter;
	EXTREACTIONCOUNTERWARNINGLOCK : L_IE1P_ReactionCounter;
	EXTREACTIONCOUNTERFAULTLOG : L_IE1P_ReactionCounter;
	EXTREACTIONCOUNTERFAULT : L_IE1P_ReactionCounter;
	EXTSEVERITYCOUNTER : L_IE1P_SeverityCounter;
	FORWARDEDSEVERITYMM : L_IE1P_SeverityLevel;
	FORWARDEDREACTIONMM : L_IE1P_Reaction;
	FORWARDEDSEVERITYSTATUSMM : L_IE1P_SeverityStatus;
	FORWARDEDREACTIONSTATUSMM : L_IE1P_ReactionStatus;
	FORWARDEDAFFECTEDMODULEMM : L_IMHP_IModuleHandler;
	FORWARDERRORHANDLER : RTS_IEC_HANDLE;
	FORWARDMODULEHANDLER : L_IMHP_IModuleHandler;
	CHILDAFTERONLINECHANGE : L_IMHP_IModuleHandler;
	PARENTAFTERONLINECHANGE : L_IMHP_IModuleHandler;
	CHILDRELATIONSHIPAFTERONLINECHANGE : L_IMHP_RelationshipID;
	PARENTRELATIONSHIPAFTERONLINECHANGE : L_IMHP_RelationshipID;
	XUPDATEACTIVESTATUSAFTERONLINECHANGE : BOOL;
	XUPDATEMODULENAMEAFTERONLINECHANGE : BOOL;
	XFORWARDSEVERITYTOPARENT : BOOL := TRUE;
	XLAYERWASSET : BOOL := FALSE;
	XFORWARDSEVERITIES : BOOL;
	XFORWARDSEVERITIESASEXTERN : BOOL;
	XMODULEREGISTERATONLINECHANGEBUSY : BOOL := FALSE;
	XLLMAVAILABLE : BOOL := FALSE;
	XLAMAVAILABLE : BOOL := FALSE;
	MAXSERVICES : UINT := 5;
	MAXCHILD : UINT := 18;
	COMPACTIVEDEFAULT : BOOL;
	COMPNAME : STRING;
	COMPTYPE : L_IMHP_ComponentType;
	DEFAULTRELATIONSHIP : L_IMHP_RelationshipID;
	ERRORHANDLE : RTS_IEC_HANDLE;
	FORWARDLOGENTRYENABLED : BOOL;
	FORWARDSEVERITYTOPARENT : BOOL;
	GETMODULEHANDLERFB : POINTER TO BYTE;
	INSTANCEID : DWORD;
	LAYER : L_IMHP_Layer;
	MODULEHANDLE : RTS_IEC_HANDLE;
	REGISTERONAPPLICATIONVIEW : BOOL;
	REGISTERSERVICELEM : BOOL;
	REGISTRATIONBUSY : BOOL;
	SUBCOMPTYPE : DWORD;
	SUSPENDREGISTRATION : BOOL;
	TEXTREFID : WORD;
	USELEM : BOOL;
	USELLM : BOOL;
END_VAR
END_FUNCTION_BLOCK

METHOD SETDEVICECONNECTOR
VAR_INPUT
	PCONNECTOR : POINTER TO IoConfigConnector;
END_VAR
END_METHOD

METHOD SETLICENSEINFO
VAR_INPUT
	UDIAPPLICATIONCREDIT : DWORD := 0;
	ELICENSECLASS : L_IMHP_LM_LicensClass;
	UDILICENSECLASSNUMBER : DWORD := 0;
END_VAR
END_METHOD

METHOD SETLICENSEINFOSTR
VAR_INPUT
	SLICINFO : STRING;
END_VAR
END_METHOD

METHOD SYNCSEVERITYANDREACTIONCOUNTER
VAR_INPUT
	XHANDLEASFORWARDEDSEVERITY : BOOL;
END_VAR
VAR_IN_OUT
	SEVERITYCOUNTER_CHILD : L_IE1P_SeverityCounter;
	REACTIONCOUNTER_CHILD : L_IE1P_ReactionCounter;
	REACTIONCOUNTERWARNING_CHILD : L_IE1P_ReactionCounter;
	REACTIONCOUNTERINFORMATION_CHILD : L_IE1P_ReactionCounter;
	REACTIONCOUNTERWARNINGLOCK_CHILD : L_IE1P_ReactionCounter;
	REACTIONCOUNTERFAULTLOG_CHILD : L_IE1P_ReactionCounter;
	REACTIONCOUNTERFAULT_CHILD : L_IE1P_ReactionCounter;
END_VAR
END_METHOD

METHOD UPDATEINFOID
END_METHOD

METHOD EVENTCALLBACK : UDINT
VAR_INPUT
	PEVENTPARAM : POINTER TO EventParam;
END_VAR
END_METHOD

METHOD REGISTEREVENT
VAR_INPUT
	XONLYCALLBACKFUNCTION : BOOL;
END_VAR
END_METHOD

METHOD UNREGISTEREVENT
VAR_INPUT
	XONLYCALLBACKFUNCTION : BOOL;
END_VAR
END_METHOD

METHOD DOREGISTER
END_METHOD

METHOD UPDATEDEPENDENCIES
END_METHOD

METHOD GETSTRINGS
END_METHOD

METHOD REGISTERONLMH : BOOL
END_METHOD

METHOD AFTERGLOBALINIT
END_METHOD

METHOD FB_REINIT : BOOL
END_METHOD

METHOD FB_EXIT : BOOL
VAR_INPUT
	BINCOPYCODE : BOOL;
END_VAR
END_METHOD

METHOD FB_INIT : BOOL
VAR_INPUT
	BINITRETAINS : BOOL;
	BINCOPYCODE : BOOL;
END_VAR
END_METHOD

METHOD ACTIVATEAPPCREDITS : BOOL
VAR_INPUT
	XACTIVATE : BOOL;
END_VAR
END_METHOD

METHOD ADDAPPCREDIT
VAR_INPUT
	CREDIT : UDINT;
END_VAR
END_METHOD

METHOD CHECKERRORRESETOCCURED : BOOL
VAR_IN_OUT
	RESETTIME : SYSTIME;
END_VAR
END_METHOD

METHOD CHECKERRORRESETTRIGGER : BOOL
VAR_IN_OUT
	LASTTRIGGERTIME : TIME;
END_VAR
END_METHOD

METHOD CLEARREACTION
VAR_INPUT
	EREACTION : L_IE1P_Reaction;
	DIREACTIONCOUNT : DINT;
END_VAR
VAR_IN_OUT
	REACTIONCOUNTER : L_IE1P_ReactionCounter;
	REACTIONCOUNTERSEVERITY : L_IE1P_ReactionCounter;
END_VAR
END_METHOD

METHOD CLEARSEVERITYANDREACTION
VAR_INPUT
	ESEVERITY : USINT;
	DISEVERITYCOUNT : DINT;
	EREACTION : WORD;
	DIREACTIONCOUNT : DINT;
	XHANDLEASFORWARDEDSEVERITY : BOOL;
END_VAR
END_METHOD

METHOD FORWARDLOGENTRYCLEAR
VAR_INPUT
	WERRORID : WORD;
	WTEXTREFID : WORD;
END_VAR
END_METHOD

METHOD FORWARDLOGENTRYNOTIFY
VAR_INPUT
	WERRORID : WORD;
	WTEXTREFID : WORD;
	SEVERITY : USINT;
	REACTION : UINT;
	PRIORITY : USINT;
	GROUP : USINT;
END_VAR
END_METHOD

METHOD FORWARDSEVERITYSUBMODULES
VAR_INPUT
	XENABLE : BOOL;
END_VAR
END_METHOD

METHOD GETREACTION : L_IE1P_Reaction
VAR_INPUT
	REACTIONCOUNTER : L_IE1P_ReactionCounter;
END_VAR
END_METHOD

METHOD GETSEVERITY2
VAR_INPUT
	XINCLUDECHILDREN : BOOL;
	XDISABLESUBMODULES : BOOL := FALSE;
	XDISABLEINTERNALCHILDS : BOOL := FALSE;
	XINCLUDEOWNMODULE : BOOL := TRUE;
	XINCLUDEEXTMODULE : BOOL := TRUE;
	PSEVERITYSTATUS : POINTER TO BYTE;
	PREACTIONSTATUS : POINTER TO BYTE;
END_VAR
VAR_OUTPUT
	EHIGHESTSEVERITY : USINT;
	EHIGHESTREACTION : WORD;
	AFFECTEDMODULE : L_IMHP_IModuleHandler;
END_VAR
END_METHOD

METHOD GETSEVERITYCHILD
VAR_INPUT
	WCHILD : WORD;
END_VAR
VAR_OUTPUT
	EHIGHESTSEVERITY : USINT;
	EHIGHESTREACTION : WORD;
	AFFECTEDMODULE : L_IMHP_IModuleHandler;
END_VAR
END_METHOD

METHOD GETSEVERITY
VAR_INPUT
	XINCLUDECHILDREN : BOOL;
	XDISABLESUBMODULES : BOOL;
	XINCLUDEOWNMODULE : BOOL;
	XINCLUDEEXTMODULE : BOOL;
	PSEVERITYSTATUS : POINTER TO BYTE;
	PREACTIONSTATUS : POINTER TO BYTE;
END_VAR
VAR_OUTPUT
	EHIGHESTSEVERITY : USINT;
	EHIGHESTREACTION : WORD;
	AFFECTEDMODULE : L_IMHP_IModuleHandler;
END_VAR
END_METHOD

METHOD READACTUALERRORCODE
VAR_OUTPUT
	ESEVERITY : USINT;
	EREACTION : WORD;
	DWERRORCODE : DWORD;
END_VAR
END_METHOD

METHOD RESETCHILDERROR
END_METHOD

METHOD RESETCHILDERROR2
VAR_INPUT
	PERRORLIST : POINTER TO RTS_IEC_HANDLE;
	PWCOUNT : POINTER TO WORD;
	MAXCOUNT : WORD;
END_VAR
END_METHOD

METHOD SETERRORRESETTRIGGER
END_METHOD

METHOD SETPARENT
VAR_INPUT
	MODULEHANDLERPARENT : L_IMHP_IModuleHandler;
	RELATIONSHIP : L_IMHP_RelationshipID := L_IMHP_RelationshipID.ApplicationView;
END_VAR
END_METHOD

METHOD UPDATEACTIVESTATUS
VAR_INPUT
	XACTIVE : BOOL;
END_VAR
END_METHOD

METHOD UPDATECOMMPATH
VAR_INPUT
	SPATH : STRING(199);
END_VAR
END_METHOD

METHOD UPDATECOMPONENTTYPE
VAR_INPUT
	ECOMPTYPE : L_IMHP_ComponentType;
END_VAR
END_METHOD

METHOD UPDATEREACTION
VAR_INPUT
	EREACTION : L_IE1P_Reaction;
END_VAR
VAR_IN_OUT
	REACTIONCOUNTER : L_IE1P_ReactionCounter;
	REACTIONCOUNTERSEVERITY : L_IE1P_ReactionCounter;
END_VAR
END_METHOD

METHOD UPDATESEVERITYANDREACTION
VAR_INPUT
	ESEVERITY : USINT;
	EREACTION : WORD;
	XHANDLEASFORWARDEDSEVERITY : BOOL;
END_VAR
END_METHOD

METHOD ADDCHILD
VAR_INPUT
	MODULEHANDLERCHILD : L_IMHP_IModuleHandler;
	RELATIONSHIP : L_IMHP_RelationshipID := L_IMHP_RelationshipID.ApplicationView;
END_VAR
END_METHOD

METHOD GETCHILD : L_IMHP_IModuleHandler
VAR_INPUT
	WNBR : WORD;
END_VAR
END_METHOD

METHOD REMOVECHILD
VAR_INPUT
	MODULEHANDLERCHILD : L_IMHP_IModuleHandler;
END_VAR
END_METHOD

METHOD SETCHILDFORDELAYEDREGISTRATION
VAR_INPUT
	MODULEHANDLERCHILD : L_IMHP_IModuleHandler;
	RELATIONSHIP : L_IMHP_RelationshipID := L_IMHP_RelationshipID.ApplicationView;
END_VAR
END_METHOD

METHOD GETCOMMPATH
VAR_IN_OUT
	SCOMMPATH : STRING(199);
END_VAR
END_METHOD

METHOD GETCOMPTYPE : L_IMHP_ComponentType
END_METHOD

METHOD GETDEVICECONNECTOR : POINTER TO IoConfigConnector
END_METHOD

METHOD GETMODULEINFO : BOOL
VAR_IN_OUT
	MODULEINFO : L_IMHP_ModuleInfo;
END_VAR
END_METHOD

METHOD GETMODULENAME
VAR_IN_OUT
	SNAME : STRING;
END_VAR
END_METHOD

METHOD REGISTEREDONSERVICE : BOOL
VAR_INPUT
	SERVICEID : L_IMHP_ServiceID;
END_VAR
END_METHOD

(* ---- L_IMHP_MODULEHANDLERTEMPLATE.pou ---- *)
FUNCTION_BLOCK L_IMHP_MODULEHANDLERTEMPLATE
VAR
	COMPNAME : STRING;
	ERRORHANDLE : SysTypes.RTS_IEC_HANDLE;
	FORWARDLOGENTRYENABLED : BOOL;
	FORWARDSEVERITYTOPARENT : BOOL;
	GETMODULEHANDLERFB : POINTER TO BYTE;
	INSTANCEID : DWORD;
	MODULEHANDLE : SysTypes.RTS_IEC_HANDLE;
	REGISTRATIONBUSY : BOOL;
END_VAR
END_FUNCTION_BLOCK

METHOD ACTIVATEAPPCREDITS : BOOL
VAR_INPUT
	XACTIVATE : BOOL;
END_VAR
END_METHOD

METHOD ADDAPPCREDIT
VAR_INPUT
	CREDIT : UDINT;
END_VAR
END_METHOD

METHOD ADDCHILD
VAR_INPUT
	MODULEHANDLERCHILD : L_IMHP_IModuleHandler;
	RELATIONSHIP : L_IMHP_RelationshipID := L_IMHP_RelationshipID.ApplicationView;
END_VAR
END_METHOD

METHOD CHECKERRORRESETOCCURED : BOOL
VAR_IN_OUT
	RESETTIME : SysTimeCore.SYSTIME;
END_VAR
END_METHOD

METHOD CHECKERRORRESETTRIGGER : BOOL
VAR_IN_OUT
	LASTTRIGGERTIME : TIME;
END_VAR
END_METHOD

METHOD CLEARSEVERITYANDREACTION
VAR_INPUT
	ESEVERITY : USINT;
	DISEVERITYCOUNT : DINT;
	EREACTION : WORD;
	DIREACTIONCOUNT : DINT;
	XHANDLEASFORWARDEDSEVERITY : BOOL;
END_VAR
END_METHOD

METHOD FORWARDLOGENTRYCLEAR
VAR_INPUT
	WERRORID : WORD;
	WTEXTREFID : WORD;
END_VAR
END_METHOD

METHOD FORWARDLOGENTRYNOTIFY
VAR_INPUT
	WERRORID : WORD;
	WTEXTREFID : WORD;
	SEVERITY : USINT;
	REACTION : UINT;
	PRIORITY : USINT;
	GROUP : USINT;
END_VAR
END_METHOD

METHOD FORWARDSEVERITYSUBMODULES
VAR_INPUT
	XENABLE : BOOL;
END_VAR
END_METHOD

METHOD GETCHILD : L_IMHP_IModuleHandler
VAR_INPUT
	WNBR : WORD;
END_VAR
END_METHOD

METHOD GETCOMMPATH
VAR_IN_OUT
	SCOMMPATH : STRING(199);
END_VAR
END_METHOD

METHOD GETCOMPTYPE : L_IMHP_ComponentType
END_METHOD

METHOD GETDEVICECONNECTOR : POINTER TO IoConfigConnector
END_METHOD

METHOD GETMODULEINFO : BOOL
VAR_IN_OUT
	MODULEINFO : L_IMHP_ModuleInfo;
END_VAR
END_METHOD

METHOD GETMODULENAME
VAR_IN_OUT
	SNAME : STRING;
END_VAR
END_METHOD

METHOD GETSEVERITY
VAR_INPUT
	XINCLUDECHILDREN : BOOL;
	XDISABLESUBMODULES : BOOL;
	XINCLUDEOWNMODULE : BOOL;
	XINCLUDEEXTMODULE : BOOL;
	PSEVERITYSTATUS : POINTER TO BYTE;
	PREACTIONSTATUS : POINTER TO BYTE;
END_VAR
VAR_OUTPUT
	EHIGHESTSEVERITY : USINT;
	EHIGHESTREACTION : WORD;
	AFFECTEDMODULE : L_IMHP_IModuleHandler;
END_VAR
END_METHOD

METHOD GETSEVERITY2
VAR_INPUT
	XINCLUDECHILDREN : BOOL;
	XDISABLESUBMODULES : BOOL := FALSE;
	XDISABLEINTERNALCHILDS : BOOL := FALSE;
	XINCLUDEOWNMODULE : BOOL := TRUE;
	XINCLUDEEXTMODULE : BOOL := TRUE;
	PSEVERITYSTATUS : POINTER TO BYTE;
	PREACTIONSTATUS : POINTER TO BYTE;
END_VAR
VAR_OUTPUT
	EHIGHESTSEVERITY : USINT;
	EHIGHESTREACTION : WORD;
	AFFECTEDMODULE : L_IMHP_IModuleHandler;
END_VAR
END_METHOD

METHOD GETSEVERITYCHILD
VAR_INPUT
	WCHILD : WORD;
END_VAR
VAR_OUTPUT
	EHIGHESTSEVERITY : USINT;
	EHIGHESTREACTION : WORD;
	AFFECTEDMODULE : L_IMHP_IModuleHandler;
END_VAR
END_METHOD

METHOD READACTUALERRORCODE
VAR_OUTPUT
	ESEVERITY : USINT;
	EREACTION : WORD;
	DWERRORCODE : DWORD;
END_VAR
END_METHOD

METHOD REGISTEREDONSERVICE : BOOL
VAR_INPUT
	SERVICEID : L_IMHP_ServiceID;
END_VAR
END_METHOD

METHOD REMOVECHILD
VAR_INPUT
	MODULEHANDLERCHILD : L_IMHP_IModuleHandler;
END_VAR
END_METHOD

METHOD RESETCHILDERROR
END_METHOD

METHOD RESETCHILDERROR2
VAR_INPUT
	PERRORLIST : POINTER TO RTS_IEC_HANDLE;
	PWCOUNT : POINTER TO WORD;
	MAXCOUNT : WORD;
END_VAR
END_METHOD

METHOD SETCHILDFORDELAYEDREGISTRATION
VAR_INPUT
	MODULEHANDLERCHILD : L_IMHP_IModuleHandler;
	RELATIONSHIP : L_IMHP_RelationshipID := L_IMHP_RelationshipID.ApplicationView;
END_VAR
END_METHOD

METHOD SETERRORRESETTRIGGER
END_METHOD

METHOD SETPARENT
VAR_INPUT
	MODULEHANDLERPARENT : L_IMHP_IModuleHandler;
	RELATIONSHIP : L_IMHP_RelationshipID := L_IMHP_RelationshipID.ApplicationView;
END_VAR
END_METHOD

METHOD SYNCSEVERITYANDREACTIONCOUNTER
VAR_INPUT
	XHANDLEASFORWARDEDSEVERITY : BOOL;
END_VAR
VAR_IN_OUT
	SEVERITYCOUNTER_CHILD : L_IE1P_SeverityCounter;
	REACTIONCOUNTER_CHILD : L_IE1P_ReactionCounter;
	REACTIONCOUNTERWARNING_CHILD : L_IE1P_ReactionCounter;
	REACTIONCOUNTERINFORMATION_CHILD : L_IE1P_ReactionCounter;
	REACTIONCOUNTERWARNINGLOCK_CHILD : L_IE1P_ReactionCounter;
	REACTIONCOUNTERFAULTLOG_CHILD : L_IE1P_ReactionCounter;
	REACTIONCOUNTERFAULT_CHILD : L_IE1P_ReactionCounter;
END_VAR
END_METHOD

METHOD UPDATEACTIVESTATUS
VAR_INPUT
	XACTIVE : BOOL;
END_VAR
END_METHOD

METHOD UPDATESEVERITYANDREACTION
VAR_INPUT
	ESEVERITY : USINT;
	EREACTION : WORD;
	XHANDLEASFORWARDEDSEVERITY : BOOL;
END_VAR
END_METHOD

(* ---- L_IMHP_WRITECOMPONENTLIST.pou ---- *)
FUNCTION_BLOCK L_IMHP_WRITECOMPONENTLIST
VAR_INPUT
	XEXECUTE : BOOL;
	SFILENAME : STRING := '';
END_VAR
VAR_OUTPUT
	XBUSY : BOOL;
	XDONE : BOOL;
	XERROR : BOOL;
	EERRORID : L_IE1P_Error;
END_VAR
VAR
	XEXECUTEOLD : BOOL;
	XREADY_INT : BOOL;
	XRESETOUTPUT : BOOL;
	SFILE_INT : STRING := '';
END_VAR
END_FUNCTION_BLOCK

METHOD ABORT : UDINT
END_METHOD

METHOD EXECUTE : UDINT
END_METHOD
